Fanuc KAREL source: KA00062.KL

PROGRAM KA00062
%NOLOCKGROUP
VAR
  SRC: XYZWPR
  DST: REAL
BEGIN
  SRC.X = 1.0
  DST = SRC
END KA00062
